// TIA Portal V21 export
VAR_GLOBAL   // PLC tag table "ConstantReady"
END_VAR
VAR_GLOBAL CONSTANT   // user constants
   SR_NO_READY : Int := 0;
   SR_READY : Int := 1;
END_VAR
